(* CODESYS project Tc3_McCollisionAvoidance.library
   TcLibraryId: Beckhoff Automation GmbH|Tc3_McCollisionAvoidance|4.0.17.0
   Company: Beckhoff Automation GmbH
   Title: Tc3_McCollisionAvoidance
   Placeholder: Tc3_McCollisionAvoidance
   Version: 4.0.17.0

Project tree, tasks and I/O mapping:
  libraries: Tc2_MC2, * (Beckhoff Automation GmbH); Tc3_Mc3Definitions, 4.0.17.0 (Beckhoff Automation GmbH)
  POUs/
    Administrative/
      function block MC_ActivateTrack [ST]: FB_init, FB_exit
      function block MC_ReadTrackPositions [ST]: FB_init, FB_exit
    Motion/
      function block MC_GearInPosCA [ST]: FB_init, FB_exit
      function block MC_HaltCA [ST]: FB_init, FB_exit
      function block MC_MoveAbsoluteCA [ST]: FB_init, FB_exit
      function block MC_MoveRelativeCA [ST]: FB_init, FB_exit
  DUTs/
    data type MC_GAP_CONTROL_MODE
    data type MC_MASTER_SIGNAL_CORRECTION
    data type ST_GearInCAOptions
    data type ST_GearInPosCAOptions
    data type ST_HaltCAOptions
    data type ST_MoveAbsoluteCAOptions
    data type ST_MoveRelativeCAOptions
  Version/
    global variables Global_Version
*)

// DUTs/MC_GAP_CONTROL_MODE
{attribute 'TcIecLibraryType'}
{attribute 'Namespace' := 'Tc3_McCollisionAvoidance'}
TYPE MC_GAP_CONTROL_MODE : (mcGapControlModeGroupDefault:=0, mcGapControlModeStandard:=1, mcGapControlModeFast:=2, mcGapControlModeNone:=3) UDINT;
END_TYPE

// DUTs/MC_MASTER_SIGNAL_CORRECTION
{attribute 'TcIecLibraryType'}
{attribute 'Namespace' := 'Tc3_McCollisionAvoidance'}
TYPE MC_MASTER_SIGNAL_CORRECTION : (mcMasterSignalCorrectionAuto:=0, mcMasterSignalCorrectionNone:=1) WORD;
END_TYPE

// DUTs/ST_GearInCAOptions
{attribute 'TcIecLibraryType'}
{attribute 'Namespace' := 'Tc3_McCollisionAvoidance'}
{attribute 'hide'}
TYPE ST_GearInCAOptions : 
	STRUCT
		{attribute 'GUID' := '78514C06-BDC7-4ADC-BF69-DC460C40C527'}
		{attribute 'Namespace' := 'Tc3_McCollisionAvoidance'}
		GapControlMode : MC_GAP_CONTROL_MODE := 0;
	END_STRUCT
END_TYPE

// DUTs/ST_GearInPosCAOptions
(* The Options can be set to specialize the synchronization profile of the slave further. *)
{attribute 'TcIecLibraryType'}
{attribute 'Namespace' := 'Tc3_McCollisionAvoidance'}
TYPE ST_GearInPosCAOptions : 
	STRUCT
		(* Maximal slave axis velocity after the slave has become synchronous for the first time. The velocity is limited by the maximum slave axis velocity. If no value is entered, the default value is used (see CA-Group Parameter GearInPosAfterSyncDynamics). *)
		{attribute 'GUID' := '0100FF8A-3F83-4535-990A-614CFBA4DA63'}
		{attribute 'Namespace' := 'MC'}
		AfterSyncVelocity : MC.MC_LREAL := MC_DEFAULT;
		(* Maximal slave axis acceleration after the slave has become synchronous for the first time. The acceleration is limited by the maximum slave axis acceleration. If no value is entered, the default value is used (see CA-Group Parameter GearInPosAfterSyncDynamics). *)
		{attribute 'GUID' := '0100FF8A-3F83-4535-990A-614CFBA4DA63'}
		{attribute 'Namespace' := 'MC'}
		AfterSyncAcceleration : MC.MC_LREAL := MC_DEFAULT;
		(* Maximal slave axis deceleration after the slave has become synchronous for the first time. The deceleration is limited by the maximum slave axis deceleration. If no value is entered, the default value is used (see CA-Group Parameter GearInPosAfterSyncDynamics). *)
		{attribute 'GUID' := '0100FF8A-3F83-4535-990A-614CFBA4DA63'}
		{attribute 'Namespace' := 'MC'}
		AfterSyncDeceleration : MC.MC_LREAL := MC_DEFAULT;
		(* Maximal slave axis jerk after the slave has become synchronous for the first time. The jerk is not limited by other jerk values (an axis maximum jerk cannot be configured). If no value is entered, the default value is used (see CA-Group Parameter GearInPosAfterSyncDynamics). *)
		{attribute 'GUID' := '0100FF8A-3F83-4535-990A-614CFBA4DA63'}
		{attribute 'Namespace' := 'MC'}
		AfterSyncJerk : MC.MC_LREAL := MC_DEFAULT;
		(* If set to FALSE, the slave velocity during the synchronization phase is always larger or equal to the master velocity. *)
		MasterVelocityUndershootAllowed : BOOL := TRUE;
		(* If set to FALSE, the slave velocity during the synchronization phase is always smaller or equal to the master velocity. *)
		MasterVelocityOvershootAllowed : BOOL := TRUE;
		 {attribute 'hide'}
		_reserved1 : ARRAY [1..6] OF USINT;
		(* Absolute minimal position of the slave during the synchronization phase. This option has effect only on the synchronization profile and has no effect once the slave is InSync. *)
		{attribute 'GUID' := '0100FF8A-3F83-4535-990A-614CFBA4DA63'}
		{attribute 'Namespace' := 'MC'}
		MinimalSlavePosition : MC.MC_LREAL := MC_IGNORE;
		(* If set to FALSE, the slave is not allowed to move in the opposite direction. *)
		DirectionReversalAllowed : BOOL := TRUE;
		(* If set to TRUE, the movement of the master is impressed on the synchronization profile of the slave, the synchronization profile is not recalculated if the master velocity changes. *)
		OverrideSlaveDynamicRestrictions : BOOL := FALSE;
		 {attribute 'hide'}
		_reserved2 : UINT;
		{attribute 'GUID' := '78514C06-BDC7-4ADC-BF69-DC460C40C527'}
		{attribute 'Namespace' := 'Tc3_McCollisionAvoidance'}
		GapControlMode : MC_GAP_CONTROL_MODE := mcGapControlModeGroupDefault;
		{attribute 'GUID' := '18071995-0000-0000-0000-00000000000F'}
		SlaveSyncPositionReferenceSystem : GLOBAL.OTCID := 0;
		{attribute 'GUID' := '18071995-0000-0000-0000-00000000000F'}
		DynamicsReferenceSystem : GLOBAL.OTCID := 0;
		(* Specifies whether and how the input from the master is corrected before being processed further by the GearInPosCA. *)
		{attribute 'GUID' := '78E5C1CC-ED57-44D7-A525-6A459863ECC4'}
		{attribute 'Namespace' := 'Tc3_McCollisionAvoidance'}
		MasterSignalCorrection : MC_MASTER_SIGNAL_CORRECTION := mcMasterSignalCorrectionAuto;
		 {attribute 'hide'}
		_reserved3 : ARRAY [1..6] OF USINT;
	END_STRUCT
END_TYPE

// DUTs/ST_HaltCAOptions
{attribute 'TcIecLibraryType'}
{attribute 'Namespace' := 'Tc3_McCollisionAvoidance'}
TYPE ST_HaltCAOptions : 
	STRUCT
		{attribute 'GUID' := '78514C06-BDC7-4ADC-BF69-DC460C40C527'}
		{attribute 'Namespace' := 'Tc3_McCollisionAvoidance'}
		GapControlMode : MC_GAP_CONTROL_MODE := 0;
		{attribute 'GUID' := '18071995-0000-0000-0000-00000000000F'}
		DynamicsReferenceSystem : GLOBAL.OTCID := 0;
	END_STRUCT
END_TYPE

// DUTs/ST_MoveAbsoluteCAOptions
{attribute 'TcIecLibraryType'}
{attribute 'Namespace' := 'Tc3_McCollisionAvoidance'}
TYPE ST_MoveAbsoluteCAOptions : 
	STRUCT
		{attribute 'GUID' := '78514C06-BDC7-4ADC-BF69-DC460C40C527'}
		{attribute 'Namespace' := 'Tc3_McCollisionAvoidance'}
		GapControlMode : MC_GAP_CONTROL_MODE := 0;
		{attribute 'GUID' := '18071995-0000-0000-0000-00000000000F'}
		PositionReferenceSystem : GLOBAL.OTCID := 0;
		{attribute 'GUID' := '18071995-0000-0000-0000-00000000000F'}
		DynamicsReferenceSystem : GLOBAL.OTCID := 0;
		AdditionalTurns : UDINT := 0;
	END_STRUCT
END_TYPE

// DUTs/ST_MoveRelativeCAOptions
{attribute 'TcIecLibraryType'}
{attribute 'Namespace' := 'Tc3_McCollisionAvoidance'}
TYPE ST_MoveRelativeCAOptions : 
	STRUCT
		{attribute 'GUID' := '78514C06-BDC7-4ADC-BF69-DC460C40C527'}
		{attribute 'Namespace' := 'Tc3_McCollisionAvoidance'}
		GapControlMode : MC_GAP_CONTROL_MODE := 0;
		{attribute 'GUID' := '18071995-0000-0000-0000-00000000000F'}
		PositionReferenceSystem : GLOBAL.OTCID := 0;
		{attribute 'GUID' := '18071995-0000-0000-0000-00000000000F'}
		DynamicsReferenceSystem : GLOBAL.OTCID := 0;
	END_STRUCT
END_TYPE

// Version/Global_Version
{attribute 'TcGenerated'}
// This function has been automatically generated from the project information.
VAR_GLOBAL CONSTANT
	{attribute 'const_non_replaced'}
	{attribute 'linkalways'}
	stLibVersion_Tc3_McCollisionAvoidance : ST_LibVersion := (iMajor := 4, iMinor := 0, iBuild := 17, iRevision := 0, nFlags := 0, sVersion := '4.0.17.0');
	{attribute 'const_non_replaced'}
	{attribute 'linkalways'}
	sLibraryId_Tc3_McCollisionAvoidance : String := 'Beckhoff Automation GmbH|Tc3_McCollisionAvoidance|4.0.17.0';
END_VAR

// POUs/Administrative/MC_ActivateTrack

{attribute 'c++_compatible'}
{attribute 'external_name' := 'MC_ActivateTrack_GUID_16BDB9B2_49D5_B836_DCE1_EF3AE1041409'}
{attribute 'TcIecLibraryType'}
{attribute 'hide_all_locals'}
FUNCTION_BLOCK MC_ActivateTrack
VAR_IN_OUT
	{attribute 'GUID' := '796382E2-8BB1-4613-AF21-647CD1FFE3C7'}
	{attribute 'Namespace' := 'Tc2_MC2'}
	Axis : Tc2_MC2.AXIS_REF;
END_VAR
VAR_INPUT
	Execute : BOOL;
END_VAR
VAR
	 {attribute 'hide'}
	_reserved1 : ARRAY [1..3] OF USINT;
END_VAR
VAR_INPUT
	{attribute 'GUID' := '18071995-0000-0000-0000-00000000000F'}
	TrackId : GLOBAL.OTCID;
END_VAR
VAR_OUTPUT
	Done : BOOL;
	Busy : BOOL;
	Error : BOOL;
END_VAR
VAR
	 {attribute 'hide'}
	_reserved2 : USINT;
END_VAR
VAR_OUTPUT
	ErrorId : UDINT;
END_VAR
VAR
	InternalFBState : ARRAY [1..16] OF ULINT;
END_VAR

{attribute 'TcTypeSystem'}

(* Internal method *)
{attribute 'hide'}
METHOD FB_init : BOOL
VAR_INPUT
	(*  if TRUE, the retain variables are initialized (warm start / cold start) *)
	bInitRetains : BOOL;
	(*  if TRUE, the instance afterwards gets moved into the copy code (online change) *)
	bInCopyCode : BOOL;
END_VAR
END_METHOD

{attribute 'TcTypeSystem'}

(* Internal method *)
{attribute 'hide'}
METHOD FB_exit : BOOL
VAR_INPUT
	(*  if TRUE, the exit method is called for exiting an instance that is copied afterwards (online change). *)
	bInCopyCode : BOOL;
END_VAR
END_METHOD

END_FUNCTION_BLOCK

// POUs/Administrative/MC_ReadTrackPositions

{attribute 'c++_compatible'}
{attribute 'external_name' := 'MC_ReadTrackPositions_GUID_6301CB2E_D947_B3B3_C688_21B41CDC4233'}
{attribute 'TcIecLibraryType'}
{attribute 'hide_all_locals'}
FUNCTION_BLOCK MC_ReadTrackPositions
VAR_IN_OUT
	{attribute 'GUID' := '796382E2-8BB1-4613-AF21-647CD1FFE3C7'}
	{attribute 'Namespace' := 'Tc2_MC2'}
	Axis : Tc2_MC2.AXIS_REF;
END_VAR
VAR_INPUT
	Enable : BOOL;
END_VAR
VAR_OUTPUT
	Valid : BOOL;
	Busy : BOOL;
END_VAR
VAR
	 {attribute 'hide'}
	_reserved1 : ARRAY [1..5] OF USINT;
END_VAR
VAR_OUTPUT
	{attribute 'GUID' := '0100FF8A-3F83-4535-990A-614CFBA4DA63'}
	{attribute 'Namespace' := 'MC'}
	TrackPosition : MC.MC_LREAL;
	{attribute 'GUID' := '18071995-0000-0000-0000-00000000000F'}
	TrackId : GLOBAL.OTCID;
END_VAR
VAR
	 {attribute 'hide'}
	_reserved2 : UDINT;
END_VAR
VAR_OUTPUT
	{attribute 'GUID' := '0100FF8A-3F83-4535-990A-614CFBA4DA63'}
	{attribute 'Namespace' := 'MC'}
	PartPosition : MC.MC_LREAL;
	{attribute 'GUID' := '18071995-0000-0000-0000-00000000000F'}
	PartId : GLOBAL.OTCID;
	Error : BOOL;
END_VAR
VAR
	 {attribute 'hide'}
	_reserved3 : ARRAY [1..3] OF USINT;
END_VAR
VAR_OUTPUT
	ErrorId : UDINT;
END_VAR
VAR
	 {attribute 'hide'}
	_reserved4 : UINT_0_32;
	{attribute 'GUID' := '18071995-0000-0000-0000-000000000018'}
	spAxis : GLOBAL.PVOID;
END_VAR

{attribute 'TcTypeSystem'}

(* Internal method *)
{attribute 'hide'}
METHOD FB_init : BOOL
VAR_INPUT
	(*  if TRUE, the retain variables are initialized (warm start / cold start) *)
	bInitRetains : BOOL;
	(*  if TRUE, the instance afterwards gets moved into the copy code (online change) *)
	bInCopyCode : BOOL;
END_VAR
END_METHOD

{attribute 'TcTypeSystem'}

(* Internal method *)
{attribute 'hide'}
METHOD FB_exit : BOOL
VAR_INPUT
	(*  if TRUE, the exit method is called for exiting an instance that is copied afterwards (online change). *)
	bInCopyCode : BOOL;
END_VAR
END_METHOD

END_FUNCTION_BLOCK

// POUs/Motion/MC_GearInPosCA

{attribute 'c++_compatible'}
{attribute 'external_name' := 'MC_GearInPosCA_GUID_C547485E_0AE1_B9F5_E0E1_50D3FC3C0A2C'}
{attribute 'TcIecLibraryType'}
{attribute 'hide_all_locals'}
FUNCTION_BLOCK MC_GearInPosCA
VAR_IN_OUT
	{attribute 'GUID' := '796382E2-8BB1-4613-AF21-647CD1FFE3C7'}
	{attribute 'Namespace' := 'Tc2_MC2'}
	Master : Tc2_MC2.AXIS_REF;
	{attribute 'GUID' := '796382E2-8BB1-4613-AF21-647CD1FFE3C7'}
	{attribute 'Namespace' := 'Tc2_MC2'}
	Slave : Tc2_MC2.AXIS_REF;
END_VAR
VAR_INPUT
	Execute : BOOL;
	ContinuousUpdate : BOOL;
END_VAR
VAR
	 {attribute 'hide'}
	_reserved1 : UINT_16_48;
END_VAR
VAR_INPUT
	{attribute 'GUID' := '0100FF8A-3F83-4535-990A-614CFBA4DA63'}
	{attribute 'Namespace' := 'MC'}
	RatioNumerator : MC.MC_LREAL;
	RatioDenumerator : UINT;
END_VAR
VAR
	 {attribute 'hide'}
	_reserved2 : ARRAY [1..6] OF USINT;
END_VAR
VAR_INPUT
	{attribute 'GUID' := '0100FF8A-3F83-4535-990A-614CFBA4DA63'}
	{attribute 'Namespace' := 'MC'}
	MasterSyncPosition : MC.MC_LREAL;
	{attribute 'GUID' := '0100FF8A-3F83-4535-990A-614CFBA4DA63'}
	{attribute 'Namespace' := 'MC'}
	SlaveSyncPosition : MC.MC_LREAL;
	{attribute 'Namespace' := 'Tc3_Mc3Definitions'}
	SyncStrategy : Tc3_Mc3Definitions.MC_SYNC_STRATEGY;
	{attribute 'Namespace' := 'Tc3_Mc3Definitions'}
	SyncMode : Tc3_Mc3Definitions.MC_SYNC_MODE;
END_VAR
VAR
	 {attribute 'hide'}
	_reserved3 : UDINT;
END_VAR
VAR_INPUT
	{attribute 'GUID' := '0100FF8A-3F83-4535-990A-614CFBA4DA63'}
	{attribute 'Namespace' := 'MC'}
	MasterStartDistance : MC.MC_LREAL;
	{attribute 'GUID' := '0100FF8A-3F83-4535-990A-614CFBA4DA63'}
	{attribute 'Namespace' := 'MC'}
	Velocity : MC.MC_LREAL;
	{attribute 'GUID' := '0100FF8A-3F83-4535-990A-614CFBA4DA63'}
	{attribute 'Namespace' := 'MC'}
	Acceleration : MC.MC_LREAL;
	{attribute 'GUID' := '0100FF8A-3F83-4535-990A-614CFBA4DA63'}
	{attribute 'Namespace' := 'MC'}
	Deceleration : MC.MC_LREAL;
	{attribute 'GUID' := '0100FF8A-3F83-4535-990A-614CFBA4DA63'}
	{attribute 'Namespace' := 'MC'}
	Jerk : MC.MC_LREAL;
	{attribute 'GUID' := '0100FF8A-3F83-4535-990A-614CFBA4DA63'}
	{attribute 'Namespace' := 'MC'}
	Gap : MC.MC_LREAL;
	{attribute 'Namespace' := 'Tc3_Mc3Definitions'}
	BufferMode : Tc3_Mc3Definitions.MC_BUFFER_MODE;
END_VAR
VAR
	 {attribute 'hide'}
	_reserved4 : ARRAY [1..6] OF USINT;
END_VAR
VAR_INPUT
	{attribute 'GUID' := '6482574D-0732-4F97-A23A-09AD62B9B681'}
	{attribute 'Namespace' := 'Tc3_McCollisionAvoidance'}
	Options : ST_GearInPosCAOptions;
END_VAR
VAR_OUTPUT
	StartSync : BOOL;
	InSync : BOOL;
	Busy : BOOL;
	Active : BOOL;
	CommandAborted : BOOL;
	Error : BOOL;
END_VAR
VAR
	 {attribute 'hide'}
	_reserved5 : UINT;
END_VAR
VAR_OUTPUT
	ErrorId : UDINT;
END_VAR
VAR
	 {attribute 'hide'}
	_reserved6 : UDINT;
	InternalFBState : ARRAY [1..16] OF ULINT;
END_VAR

{attribute 'TcTypeSystem'}

(* Internal method *)
{attribute 'hide'}
METHOD FB_init : BOOL
VAR_INPUT
	(*  if TRUE, the retain variables are initialized (warm start / cold start) *)
	bInitRetains : BOOL;
	(*  if TRUE, the instance afterwards gets moved into the copy code (online change) *)
	bInCopyCode : BOOL;
END_VAR
END_METHOD

{attribute 'TcTypeSystem'}

(* Internal method *)
{attribute 'hide'}
METHOD FB_exit : BOOL
VAR_INPUT
	(*  if TRUE, the exit method is called for exiting an instance that is copied afterwards (online change). *)
	bInCopyCode : BOOL;
END_VAR
END_METHOD

END_FUNCTION_BLOCK

// POUs/Motion/MC_HaltCA

{attribute 'c++_compatible'}
{attribute 'external_name' := 'MC_HaltCA_GUID_AC3F6B24_69AD_B962_C838_7E76AB14E4C5'}
{attribute 'TcIecLibraryType'}
{attribute 'hide_all_locals'}
FUNCTION_BLOCK MC_HaltCA
VAR_IN_OUT
	{attribute 'GUID' := '796382E2-8BB1-4613-AF21-647CD1FFE3C7'}
	{attribute 'Namespace' := 'Tc2_MC2'}
	Axis : Tc2_MC2.AXIS_REF;
END_VAR
VAR_INPUT
	Execute : BOOL;
END_VAR
VAR
	 {attribute 'hide'}
	_reserved1 : ARRAY [1..7] OF USINT;
END_VAR
VAR_INPUT
	{attribute 'GUID' := '0100FF8A-3F83-4535-990A-614CFBA4DA63'}
	{attribute 'Namespace' := 'MC'}
	Deceleration : MC.MC_LREAL;
	{attribute 'GUID' := '0100FF8A-3F83-4535-990A-614CFBA4DA63'}
	{attribute 'Namespace' := 'MC'}
	Jerk : MC.MC_LREAL;
	{attribute 'GUID' := '0100FF8A-3F83-4535-990A-614CFBA4DA63'}
	{attribute 'Namespace' := 'MC'}
	Gap : MC.MC_LREAL;
	{attribute 'GUID' := '08EE1E90-DD03-4341-8283-229DD3F04035'}
	{attribute 'Namespace' := 'Tc3_McCollisionAvoidance'}
	Options : ST_HaltCAOptions;
END_VAR
VAR_OUTPUT
	Done : BOOL;
	Busy : BOOL;
	Active : BOOL;
	CommandAborted : BOOL;
	Error : BOOL;
END_VAR
VAR
	 {attribute 'hide'}
	_reserved2 : ARRAY [1..3] OF USINT;
END_VAR
VAR_OUTPUT
	ErrorId : UDINT;
END_VAR
VAR
	 {attribute 'hide'}
	_reserved3 : UDINT;
	InternalFBState : ARRAY [1..16] OF ULINT;
END_VAR

{attribute 'TcTypeSystem'}

(* Internal method *)
{attribute 'hide'}
METHOD FB_init : BOOL
VAR_INPUT
	(*  if TRUE, the retain variables are initialized (warm start / cold start) *)
	bInitRetains : BOOL;
	(*  if TRUE, the instance afterwards gets moved into the copy code (online change) *)
	bInCopyCode : BOOL;
END_VAR
END_METHOD

{attribute 'TcTypeSystem'}

(* Internal method *)
{attribute 'hide'}
METHOD FB_exit : BOOL
VAR_INPUT
	(*  if TRUE, the exit method is called for exiting an instance that is copied afterwards (online change). *)
	bInCopyCode : BOOL;
END_VAR
END_METHOD

END_FUNCTION_BLOCK

// POUs/Motion/MC_MoveAbsoluteCA

{attribute 'c++_compatible'}
{attribute 'external_name' := 'MC_MoveAbsoluteCA_GUID_D14738CE_75A3_B0A1_FD8C_C11E050E0E63'}
{attribute 'TcIecLibraryType'}
{attribute 'hide_all_locals'}
FUNCTION_BLOCK MC_MoveAbsoluteCA
VAR_IN_OUT
	{attribute 'GUID' := '796382E2-8BB1-4613-AF21-647CD1FFE3C7'}
	{attribute 'Namespace' := 'Tc2_MC2'}
	Axis : Tc2_MC2.AXIS_REF;
END_VAR
VAR_INPUT
	Execute : BOOL;
	ContinuousUpdate : BOOL;
END_VAR
VAR
	 {attribute 'hide'}
	_reserved1 : ARRAY [1..6] OF USINT;
END_VAR
VAR_INPUT
	{attribute 'GUID' := '0100FF8A-3F83-4535-990A-614CFBA4DA63'}
	{attribute 'Namespace' := 'MC'}
	Position : MC.MC_LREAL;
	{attribute 'GUID' := '0100FF8A-3F83-4535-990A-614CFBA4DA63'}
	{attribute 'Namespace' := 'MC'}
	Velocity : MC.MC_LREAL;
	{attribute 'GUID' := '0100FF8A-3F83-4535-990A-614CFBA4DA63'}
	{attribute 'Namespace' := 'MC'}
	Acceleration : MC.MC_LREAL;
	{attribute 'GUID' := '0100FF8A-3F83-4535-990A-614CFBA4DA63'}
	{attribute 'Namespace' := 'MC'}
	Deceleration : MC.MC_LREAL;
	{attribute 'GUID' := '0100FF8A-3F83-4535-990A-614CFBA4DA63'}
	{attribute 'Namespace' := 'MC'}
	Jerk : MC.MC_LREAL;
	{attribute 'GUID' := '0100FF8A-3F83-4535-990A-614CFBA4DA63'}
	{attribute 'Namespace' := 'MC'}
	Gap : MC.MC_LREAL;
	{attribute 'Namespace' := 'Tc3_Mc3Definitions'}
	BufferMode : Tc3_Mc3Definitions.MC_BUFFER_MODE;
	{attribute 'Namespace' := 'Tc3_Mc3Definitions'}
	Direction : Tc3_Mc3Definitions.MC_DIRECTION;
	{attribute 'GUID' := '13D285C1-E864-4752-B89D-A624CC261AFD'}
	{attribute 'Namespace' := 'Tc3_McCollisionAvoidance'}
	Options : ST_MoveAbsoluteCAOptions;
END_VAR
VAR_OUTPUT
	Done : BOOL;
	Busy : BOOL;
	Active : BOOL;
	CommandAborted : BOOL;
	Error : BOOL;
END_VAR
VAR
	 {attribute 'hide'}
	_reserved2 : ARRAY [1..3] OF USINT;
END_VAR
VAR_OUTPUT
	ErrorId : UDINT;
END_VAR
VAR
	InternalFBState : ARRAY [1..16] OF ULINT;
END_VAR

{attribute 'TcTypeSystem'}

(* Internal method *)
{attribute 'hide'}
METHOD FB_init : BOOL
VAR_INPUT
	(*  if TRUE, the retain variables are initialized (warm start / cold start) *)
	bInitRetains : BOOL;
	(*  if TRUE, the instance afterwards gets moved into the copy code (online change) *)
	bInCopyCode : BOOL;
END_VAR
END_METHOD

{attribute 'TcTypeSystem'}

(* Internal method *)
{attribute 'hide'}
METHOD FB_exit : BOOL
VAR_INPUT
	(*  if TRUE, the exit method is called for exiting an instance that is copied afterwards (online change). *)
	bInCopyCode : BOOL;
END_VAR
END_METHOD

END_FUNCTION_BLOCK

// POUs/Motion/MC_MoveRelativeCA

{attribute 'c++_compatible'}
{attribute 'external_name' := 'MC_MoveRelativeCA_GUID_745387DA_3A36_B50D_EB86_557E70158E0B'}
{attribute 'TcIecLibraryType'}
{attribute 'hide_all_locals'}
FUNCTION_BLOCK MC_MoveRelativeCA
VAR_IN_OUT
	{attribute 'GUID' := '796382E2-8BB1-4613-AF21-647CD1FFE3C7'}
	{attribute 'Namespace' := 'Tc2_MC2'}
	Axis : Tc2_MC2.AXIS_REF;
END_VAR
VAR_INPUT
	Execute : BOOL;
	ContinuousUpdate : BOOL;
END_VAR
VAR
	 {attribute 'hide'}
	_reserved1 : ARRAY [1..6] OF USINT;
END_VAR
VAR_INPUT
	{attribute 'GUID' := '0100FF8A-3F83-4535-990A-614CFBA4DA63'}
	{attribute 'Namespace' := 'MC'}
	Distance : MC.MC_LREAL;
	{attribute 'GUID' := '0100FF8A-3F83-4535-990A-614CFBA4DA63'}
	{attribute 'Namespace' := 'MC'}
	Velocity : MC.MC_LREAL;
	{attribute 'GUID' := '0100FF8A-3F83-4535-990A-614CFBA4DA63'}
	{attribute 'Namespace' := 'MC'}
	Acceleration : MC.MC_LREAL;
	{attribute 'GUID' := '0100FF8A-3F83-4535-990A-614CFBA4DA63'}
	{attribute 'Namespace' := 'MC'}
	Deceleration : MC.MC_LREAL;
	{attribute 'GUID' := '0100FF8A-3F83-4535-990A-614CFBA4DA63'}
	{attribute 'Namespace' := 'MC'}
	Jerk : MC.MC_LREAL;
	{attribute 'GUID' := '0100FF8A-3F83-4535-990A-614CFBA4DA63'}
	{attribute 'Namespace' := 'MC'}
	Gap : MC.MC_LREAL;
	{attribute 'Namespace' := 'Tc3_Mc3Definitions'}
	BufferMode : Tc3_Mc3Definitions.MC_BUFFER_MODE;
END_VAR
VAR
	 {attribute 'hide'}
	_reserved2 : UINT;
END_VAR
VAR_INPUT
	{attribute 'GUID' := '3D39C17E-DA7F-40AD-951E-99C1660F36B5'}
	{attribute 'Namespace' := 'Tc3_McCollisionAvoidance'}
	Options : ST_MoveRelativeCAOptions;
END_VAR
VAR_OUTPUT
	Done : BOOL;
	Busy : BOOL;
	Active : BOOL;
	CommandAborted : BOOL;
	Error : BOOL;
END_VAR
VAR
	 {attribute 'hide'}
	_reserved3 : ARRAY [1..3] OF USINT;
END_VAR
VAR_OUTPUT
	ErrorId : UDINT;
END_VAR
VAR
	 {attribute 'hide'}
	_reserved4 : UDINT;
	InternalFBState : ARRAY [1..16] OF ULINT;
END_VAR

{attribute 'TcTypeSystem'}

(* Internal method *)
{attribute 'hide'}
METHOD FB_init : BOOL
VAR_INPUT
	(*  if TRUE, the retain variables are initialized (warm start / cold start) *)
	bInitRetains : BOOL;
	(*  if TRUE, the instance afterwards gets moved into the copy code (online change) *)
	bInCopyCode : BOOL;
END_VAR
END_METHOD

{attribute 'TcTypeSystem'}

(* Internal method *)
{attribute 'hide'}
METHOD FB_exit : BOOL
VAR_INPUT
	(*  if TRUE, the exit method is called for exiting an instance that is copied afterwards (online change). *)
	bInCopyCode : BOOL;
END_VAR
END_METHOD

END_FUNCTION_BLOCK
